// TIA Portal V21 export
// export: Created 2026-08-21T20:18:55.5324372Z, ExportSetting None, DisplayName Totally Integrated Automation Portal, DisplayVersion V21, DisplayName STEP 7 Professional, DisplayVersion V21, DisplayName STEP 7 Safety, DisplayVersion V21, DisplayName Tech WebApplication, DisplayVersion V21, DisplayName WinCC Basic/Comfort/Advanced, DisplayVersion V21, DisplayName WinCC Professional, DisplayVersion V21, DisplayName WinCC Unified, DisplayVersion V21
TYPE "UDT_Service_Setup"
   STRUCT
      stepOrderOp : UInt;
      stepOrder { ExternalWritable := 'False'} : "UDT_Service_StepOrder";
      parameterIndexOp : UInt;
      parameterIndex { ExternalWritable := 'False'} : Byte;
   END_STRUCT;
END_TYPE
